// TIA Portal V20 export
// export: Created 2026-10-12T15:46:50.414152Z, ExportSetting WithDefaults, DisplayName Totally Integrated Automation Portal, DisplayVersion V20, DisplayName TIA Portal Openness, DisplayVersion V20, DisplayName TIA Portal Teamcenter Gateway, DisplayVersion V20, DisplayName TIA Portal Version Control Interface, DisplayVersion V20, DisplayName SINAMICS Startdrive Advanced, DisplayVersion V20 SP1 Update 2, DisplayName SINAMICS Startdrive G110M, G120, G120C, G120D, G120P, G115D, DisplayVersion V20 SP1 Update 2, DisplayName SINAMICS Startdrive G130, G150, S120, S150, SINAMICS MV, G220, S200, S210, DisplayVersion V20 SP1 Update 2, DisplayName STEP 7 Professional, DisplayVersion V20, DisplayName STEP 7 Safety, DisplayVersion V20, DisplayName WinCC Basic/Comfort/Advanced, DisplayVersion V20, DisplayName WinCC Professional, DisplayVersion V20, DisplayName WinCC Unified, DisplayVersion V20
FUNCTION "FRK_DescendantsReady" : Bool   // FC84, SCL
{ S7_Optimized_Access := 'TRUE' }
VERSION : 0.1
// stored: AutoNumber true, IsIECCheckEnabled false, SetENOAutomatically false, UDAEnableTagReadback false
   VAR_INPUT
      OwnerIndex : DInt;
   END_VAR
   VAR_TEMP
      Index : DInt;
      Parent : DInt;
      Depth : DInt;
   END_VAR
BEGIN

   #FRK_DescendantsReady := FALSE;
   IF "FRK_Registry".Fault OR #OwnerIndex < 1 OR #OwnerIndex > "FRK_Registry".Count OR "FRK_Registry".Count > 32 THEN
       RETURN;
   END_IF;
   FOR #Index := 1 TO "FRK_Registry".Count DO
       #Parent := "FRK_Registry".Rows[#Index].Parent;
       FOR #Depth := 1 TO 32 DO
           IF #Parent = #OwnerIndex THEN
               IF "FRK_Registry".Rows[#Index].Exec <> 0 THEN
                   RETURN;
               END_IF;
               EXIT;
           END_IF;
           IF #Parent = 0 THEN
               EXIT;
           END_IF;
           IF #Parent < 1 OR #Parent > "FRK_Registry".Count THEN
               RETURN;
           END_IF;
           #Parent := "FRK_Registry".Rows[#Parent].Parent;
       END_FOR;
       IF #Depth > 32 AND #Parent <> 0 THEN
           RETURN;
       END_IF;
   END_FOR;
   #FRK_DescendantsReady := TRUE;
END_FUNCTION
